Fanuc KAREL source: ka00027.KL

-- PROVISIONAL review KL for V770-1; original PC SHA256 ecf1d9a5cbef73b7de5a92310ae510402355cdb3f0758b3cf5d06c9fda734b07
-- Incomplete behavior may be omitted. Consult companion uncertainty JSON. Do not deploy.
PROGRAM KA00027
%NOLOCKGROUP
VAR
  SRC : BOOLEAN
  DST : BOOLEAN
BEGIN
  SRC = TRUE
  DST = SRC
END KA00027
